FUNCTION_BLOCK SpringMagazine (* Composite Function Block Type *)
  (* Standard: 61499-2 *)
  (* Version 0.0, 7/2/2026, template *)
  PACKAGE Main;
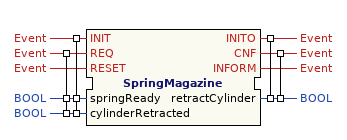
  EVENT_INPUT
    INIT WITH springReady, cylinderRetracted; (* Initialization Request *)
    REQ WITH springReady, cylinderRetracted; (* Normal Execution Request *)
    RESET;
  END_EVENT
  EVENT_OUTPUT
    INITO WITH retractCylinder; (* Initialization Confirm *)
    CNF WITH retractCylinder; (* Execution Confirmation *)
    INFORM;
  END_EVENT
  VAR_INPUT
    springReady : BOOL; (* Input event qualifier *)
    cylinderRetracted : BOOL;
  END_VAR
  VAR_OUTPUT
    retractCylinder : BOOL; (* Output event qualifier *)
  END_VAR
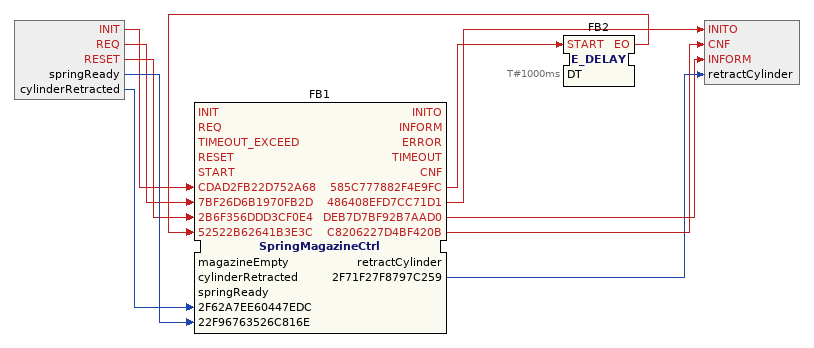
  FBS
    FB1 : SpringMagazineCtrl;
    FB2 : E_DELAY(DT := T#1000ms);
  END_FBS
  EVENT_CONNECTIONS
    INIT TO FB1.CDAD2FB22D752A68;
    REQ TO FB1.7BF26D6B1970FB2D;
    RESET TO FB1.2B6F356DDD3CF0E4;
    FB2.EO TO FB1.52522B62641B3E3C;
    FB1.585C777882F4E9FC TO FB2.START;
    FB1.486408EFD7CC71D1 TO INITO;
    FB1.DEB7D7BF92B7AAD0 TO INFORM;
    FB1.C8206227D4BF420B TO CNF;
  END_CONNECTIONS
  DATA_CONNECTIONS
    FB1.2F71F27F8797C259 TO retractCylinder;
    cylinderRetracted TO FB1.2F62A7EE60447EDC;
    springReady TO FB1.22F96763526C816E;
  END_CONNECTIONS
END_FUNCTION_BLOCK
